{region 'Documentation'}
(*!
<summary>Check that IN is greater than Minimum.</summary>
*)
{endregion}
FUNCTION_BLOCK AssertGreaterThan_USInt EXTENDS AssertionBase
VAR_INPUT
    IN : USINT; //! Actual value checked or observed by this Assertion.
    Minimum : USINT; //! Exclusive lower bound; the actual value or count must be greater.
END_VAR

SUPER^();

{region 'Documentation'}
(*!
<summary>Check that IN is greater than Minimum.</summary>
*)
{endregion}
METHOD PROTECTED Assert
VAR
    Message : STRING(GVL_Constants.MessageLength);
    MinimumText : STRING(GVL_Constants.AssertionValueLength);
    ActualText : STRING(GVL_Constants.AssertionValueLength);
END_VAR
IF NOT EvaluationActive THEN
    RETURN;
END_IF;

IF Result = E_Result.Error THEN
    RETURN;
END_IF;

IF Result = E_Result.Failed THEN
    RETURN;
END_IF;

IF IN <= Minimum THEN
    MinimumText := USINT_TO_STRING(Minimum);
    ActualText := USINT_TO_STRING(IN);
    Message := CONCAT('Assertion failed: value is not greater than minimum. Minimum = ',
        MinimumText);
    Message := CONCAT(Message, ', Actual = ');
    Message := CONCAT(Message, ActualText);
    Message := CONCAT(Message, '.');
    Fail(Message := Message);
    RETURN;
END_IF;

Pass();
END_METHOD

END_FUNCTION_BLOCK

(* stored: Version 1.1.0.1
   POU AssertGreaterThan_USInt: Id {18e0ebbf-053f-4dfb-9e1c-8695f7cf5903}, SpecialFunc None
   Folder Internal: Id {971d244c-c366-43fa-978e-91529c38d7f8}
   Method Assert: Id {700b4c23-1da0-45e7-90f7-1b6748669bbf} *)
